Staubli VAL3: savePROG.pjx

--- savePROG.pjx ---
Parameters version=s8.10.3Cs9_BS2093 stackSize=5000 millimeterUnit=true
Data file=savePROG.dtx
Type name=progItem path=Disk://source/template/progItem/progItem.pjx

--- savePROG.dtx ---
public progItem pProgItem{}
  [prod01]
    progTemplate pProgTemplate[5]
      [0]
        forItem fForItem
          [0]
            bool bIOdisable
            num nLoopValue
            string sForTRAJ
            string sIOindex
        ifItem iIfItem
          [0]
            bool bANDOR[2]
            num nSigIndex[3]
            num nSigType[3]
            num nValue[3]
        num nType
        switchItem sSwitchItem
          [0]
            bool bIOdisable
            num nSwitchValue
            string sIOValue
        string sTRAJname = "ttt"
      [1]
        forItem fForItem
          [0]
            bool bIOdisable
            num nLoopValue
            string sForTRAJ
            string sIOindex
        ifItem iIfItem
          [0]
            bool bANDOR[2]
            num nSigIndex[3]
            num nSigType[3]
            num nValue[3]
        num nType = 5
        switchItem sSwitchItem
          [0]
            bool bIOdisable = true
            num nSwitchValue
            string sIOValue = "2,工作号"
        string sTRAJname = "SWITCH"
      [2]
        forItem fForItem
          [0]
            bool bIOdisable
            num nLoopValue
            string sForTRAJ
            string sIOindex
        ifItem iIfItem
          [0]
            bool bANDOR[2]
            num nSigIndex[3]
            num nSigType[3]
            num nValue[3]
        num nType = 6
        switchItem sSwitchItem
          [0]
            bool bIOdisable
            num nSwitchValue
            string sIOValue = "prod01"
        string sTRAJname = "PROG"
      [3]
        forItem fForItem
          [0]
            bool bIOdisable
            num nLoopValue
            string sForTRAJ
            string sIOindex
        ifItem iIfItem
          [0]
            bool bANDOR[2]
            num nSigIndex[3]
            num nSigType[3]
            num nValue[3]
        num nType = 6
        switchItem sSwitchItem
          [0]
            bool bIOdisable
            num nSwitchValue = 1
            string sIOValue = "prod02"
        string sTRAJname = "PROG"
      [4]
        forItem fForItem
          [0]
            bool bIOdisable
            num nLoopValue
            string sForTRAJ
            string sIOindex
        ifItem iIfItem
          [0]
            bool bANDOR[2]
            num nSigIndex[3]
            num nSigType[3]
            num nValue[3]
        num nType = 7
        switchItem sSwitchItem
          [0]
            bool bIOdisable
            num nSwitchValue
            string sIOValue
        string sTRAJname = "ENDSWITCH"
  [prod011]
    progTemplate pProgTemplate[2]
      [0]
        forItem fForItem
          [0]
            bool bIOdisable
            num nLoopValue
            string sForTRAJ
            string sIOindex
        ifItem iIfItem
          [0]
            bool bANDOR[2]
            num nSigIndex[3]
            num nSigType[3]
            num nValue[3]
        num nType
        switchItem sSwitchItem
          [0]
            bool bIOdisable
            num nSwitchValue
            string sIOValue
        string sTRAJname = "Int"
      [1]
        forItem fForItem
          [0]
            bool bIOdisable
            num nLoopValue
            string sForTRAJ
            string sIOindex
        ifItem iIfItem
          [0]
            bool bANDOR[2]
            num nSigIndex[3]
            num nSigType[3]
            num nValue[3]
        num nType
        switchItem sSwitchItem
          [0]
            bool bIOdisable
            num nSwitchValue
            string sIOValue
        string sTRAJname = "Program011"
  [prod02]
    progTemplate pProgTemplate[2]
      [0]
        forItem fForItem
          [0]
            bool bIOdisable
            num nLoopValue
            string sForTRAJ
            string sIOindex
        ifItem iIfItem
          [0]
            bool bANDOR[2]
            num nSigIndex[3]
            num nSigType[3]
            num nValue[3]
        num nType
        switchItem sSwitchItem
          [0]
            bool bIOdisable
            num nSwitchValue
            string sIOValue
        string sTRAJname = "Int"
      [1]
        forItem fForItem
          [0]
            bool bIOdisable
            num nLoopValue
            string sForTRAJ
            string sIOindex
        ifItem iIfItem
          [0]
            bool bANDOR[2]
            num nSigIndex[3]
            num nSigType[3]
            num nValue[3]
        num nType
        switchItem sSwitchItem
          [0]
            bool bIOdisable
            num nSwitchValue
            string sIOValue
        string sTRAJname = "Program2"
  [prod03]
    progTemplate pProgTemplate[2]
      [0]
        forItem fForItem
          [0]
            bool bIOdisable
            num nLoopValue
            string sForTRAJ
            string sIOindex
        ifItem iIfItem
          [0]
            bool bANDOR[2]
            num nSigIndex[3]
            num nSigType[3]
            num nValue[3]
        num nType
        switchItem sSwitchItem
          [0]
            bool bIOdisable
            num nSwitchValue
            string sIOValue
        string sTRAJname = "Int"
      [1]
        forItem fForItem
          [0]
            bool bIOdisable
            num nLoopValue
            string sForTRAJ
            string sIOindex
        ifItem iIfItem
          [0]
            bool bANDOR[2]
            num nSigIndex[3]
            num nSigType[3]
            num nValue[3]
        num nType
        switchItem sSwitchItem
          [0]
            bool bIOdisable
            num nSwitchValue
            string sIOValue
        string sTRAJname = "Program3"
  [prod06]
    progTemplate pProgTemplate[2]
      [0]
        forItem fForItem
          [0]
            bool bIOdisable
            num nLoopValue
            string sForTRAJ
            string sIOindex
        ifItem iIfItem
          [0]
            bool bANDOR[2]
            num nSigIndex[3]
            num nSigType[3]
            num nValue[3]
        num nType
        switchItem sSwitchItem
          [0]
            bool bIOdisable
            num nSwitchValue
            string sIOValue
        string sTRAJname = "Int"
      [1]
        forItem fForItem
          [0]
            bool bIOdisable
            num nLoopValue
            string sForTRAJ
            string sIOindex
        ifItem iIfItem
          [0]
            bool bANDOR[2]
            num nSigIndex[3]
            num nSigType[3]
            num nValue[3]
        num nType
        switchItem sSwitchItem
          [0]
            bool bIOdisable
            num nSwitchValue
            string sIOValue
        string sTRAJname = "Program6"
  [prod11]
    progTemplate pProgTemplate[2]
      [0]
        forItem fForItem
          [0]
            bool bIOdisable
            num nLoopValue
            string sForTRAJ
            string sIOindex
        ifItem iIfItem
          [0]
            bool bANDOR[2]
            num nSigIndex[3]
            num nSigType[3]
            num nValue[3]
        num nType
        switchItem sSwitchItem
          [0]
            bool bIOdisable
            num nSwitchValue
            string sIOValue
        string sTRAJname = "Int"
      [1]
        forItem fForItem
          [0]
            bool bIOdisable
            num nLoopValue
            string sForTRAJ
            string sIOindex
        ifItem iIfItem
          [0]
            bool bANDOR[2]
            num nSigIndex[3]
            num nSigType[3]
            num nValue[3]
        num nType
        switchItem sSwitchItem
          [0]
            bool bIOdisable
            num nSwitchValue
            string sIOValue
        string sTRAJname = "Program11"
